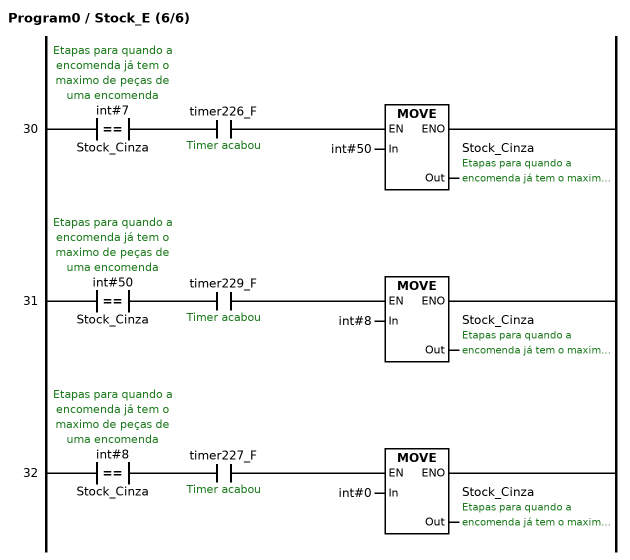
(* [picture p144: Program0 / Stock_E, rungs 30-32] *)
(* Rung 30 *)
IF (int#7 = Stock_Cinza) AND timer226_F THEN Stock_Cinza := int#50; END_IF;
(* Rung 31 *)
IF (int#50 = Stock_Cinza) AND timer229_F THEN Stock_Cinza := int#8; END_IF;
(* Rung 32 *)
IF (int#8 = Stock_Cinza) AND timer227_F THEN Stock_Cinza := int#0; END_IF;

(* Section Stock_S: ladder, written here as Structured Text *)

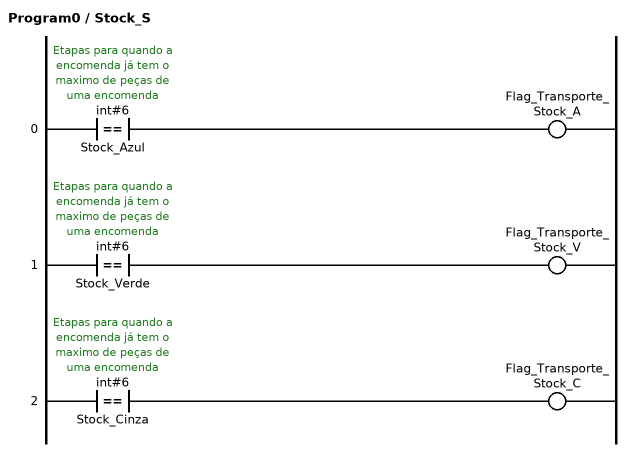
(* Rung 0 *)
Flag_Transporte_Stock_A := int#6 = Stock_Azul;
(* Rung 1 *)
Flag_Transporte_Stock_V := int#6 = Stock_Verde;
(* Rung 2 *)
Flag_Transporte_Stock_C := int#6 = Stock_Cinza;

(* Section Recolhe_Stock_E: ladder, written here as Structured Text *)

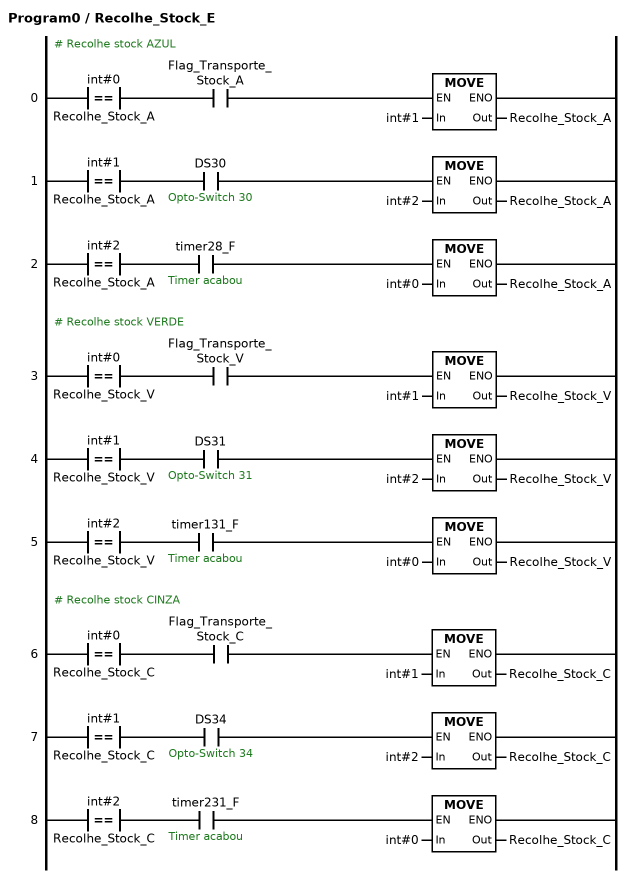
(* Rung 0: # Recolhe stock AZUL *)
IF (int#0 = Recolhe_Stock_A) AND Flag_Transporte_Stock_A THEN Recolhe_Stock_A := int#1; END_IF;
(* Rung 1 *)
IF (int#1 = Recolhe_Stock_A) AND DS30 THEN Recolhe_Stock_A := int#2; END_IF;
(* Rung 2 *)
IF (int#2 = Recolhe_Stock_A) AND timer28_F THEN Recolhe_Stock_A := int#0; END_IF;
(* Rung 3: # Recolhe stock VERDE *)
IF (int#0 = Recolhe_Stock_V) AND Flag_Transporte_Stock_V THEN Recolhe_Stock_V := int#1; END_IF;
(* Rung 4 *)
IF (int#1 = Recolhe_Stock_V) AND DS31 THEN Recolhe_Stock_V := int#2; END_IF;
(* Rung 5 *)
IF (int#2 = Recolhe_Stock_V) AND timer131_F THEN Recolhe_Stock_V := int#0; END_IF;
(* Rung 6: # Recolhe stock CINZA *)
IF (int#0 = Recolhe_Stock_C) AND Flag_Transporte_Stock_C THEN Recolhe_Stock_C := int#1; END_IF;
(* Rung 7 *)
IF (int#1 = Recolhe_Stock_C) AND DS34 THEN Recolhe_Stock_C := int#2; END_IF;
(* Rung 8 *)
IF (int#2 = Recolhe_Stock_C) AND timer231_F THEN Recolhe_Stock_C := int#0; END_IF;

(* Section Recolhe_Stock_S: ladder, written here as Structured Text *)

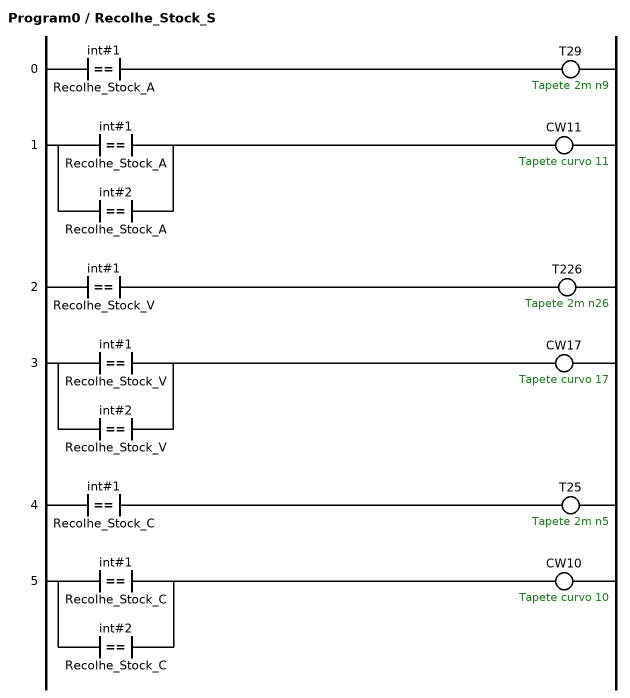
(* Rung 0 *)
T29 := int#1 = Recolhe_Stock_A;
(* Rung 1 *)
CW11 := (int#1 = Recolhe_Stock_A) OR (int#2 = Recolhe_Stock_A);
(* Rung 2 *)
T226 := int#1 = Recolhe_Stock_V;
(* Rung 3 *)
CW17 := (int#1 = Recolhe_Stock_V) OR (int#2 = Recolhe_Stock_V);
(* Rung 4 *)
T25 := int#1 = Recolhe_Stock_C;
(* Rung 5 *)
CW10 := (int#1 = Recolhe_Stock_C) OR (int#2 = Recolhe_Stock_C);

(* Section Recolha_Comum_E: ladder, written here as Structured Text *)

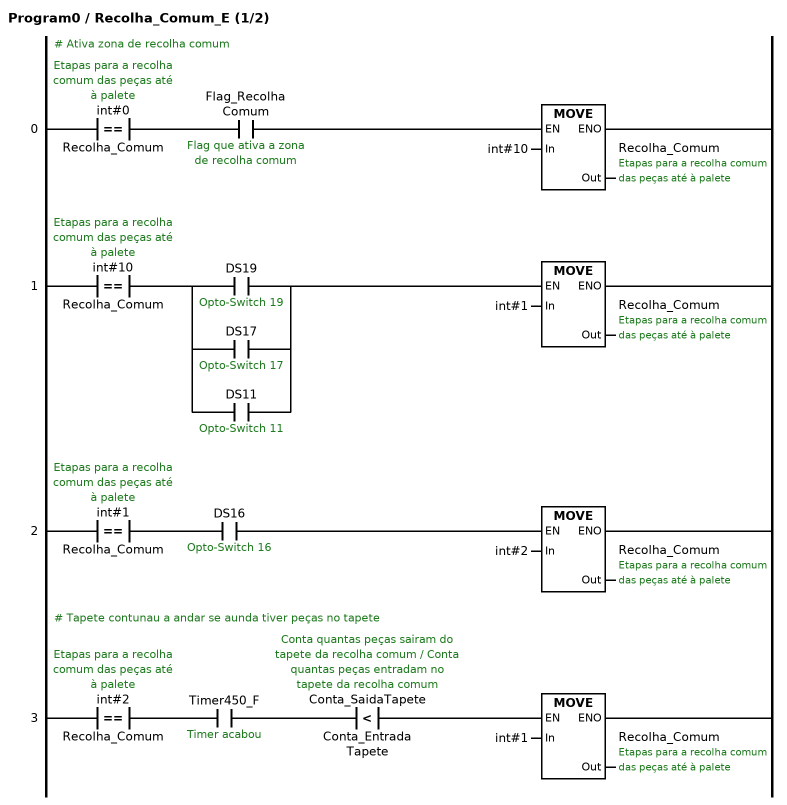
(* Rung 0: # Ativa zona de recolha comum *)
IF (int#0 = Recolha_Comum) AND Flag_RecolhaComum THEN Recolha_Comum := int#10; END_IF;
(* Rung 1 *)
IF (int#10 = Recolha_Comum) AND (DS19 OR DS17 OR DS11) THEN Recolha_Comum := int#1; END_IF;
(* Rung 2 *)
IF (int#1 = Recolha_Comum) AND DS16 THEN Recolha_Comum := int#2; END_IF;
(* Rung 3: # Tapete contunau a andar se aunda tiver peças no tapete *)
IF (int#2 = Recolha_Comum) AND Timer450_F AND (Conta_SaidaTapete < Conta_EntradaTapete) THEN
    Recolha_Comum := int#1;
END_IF;

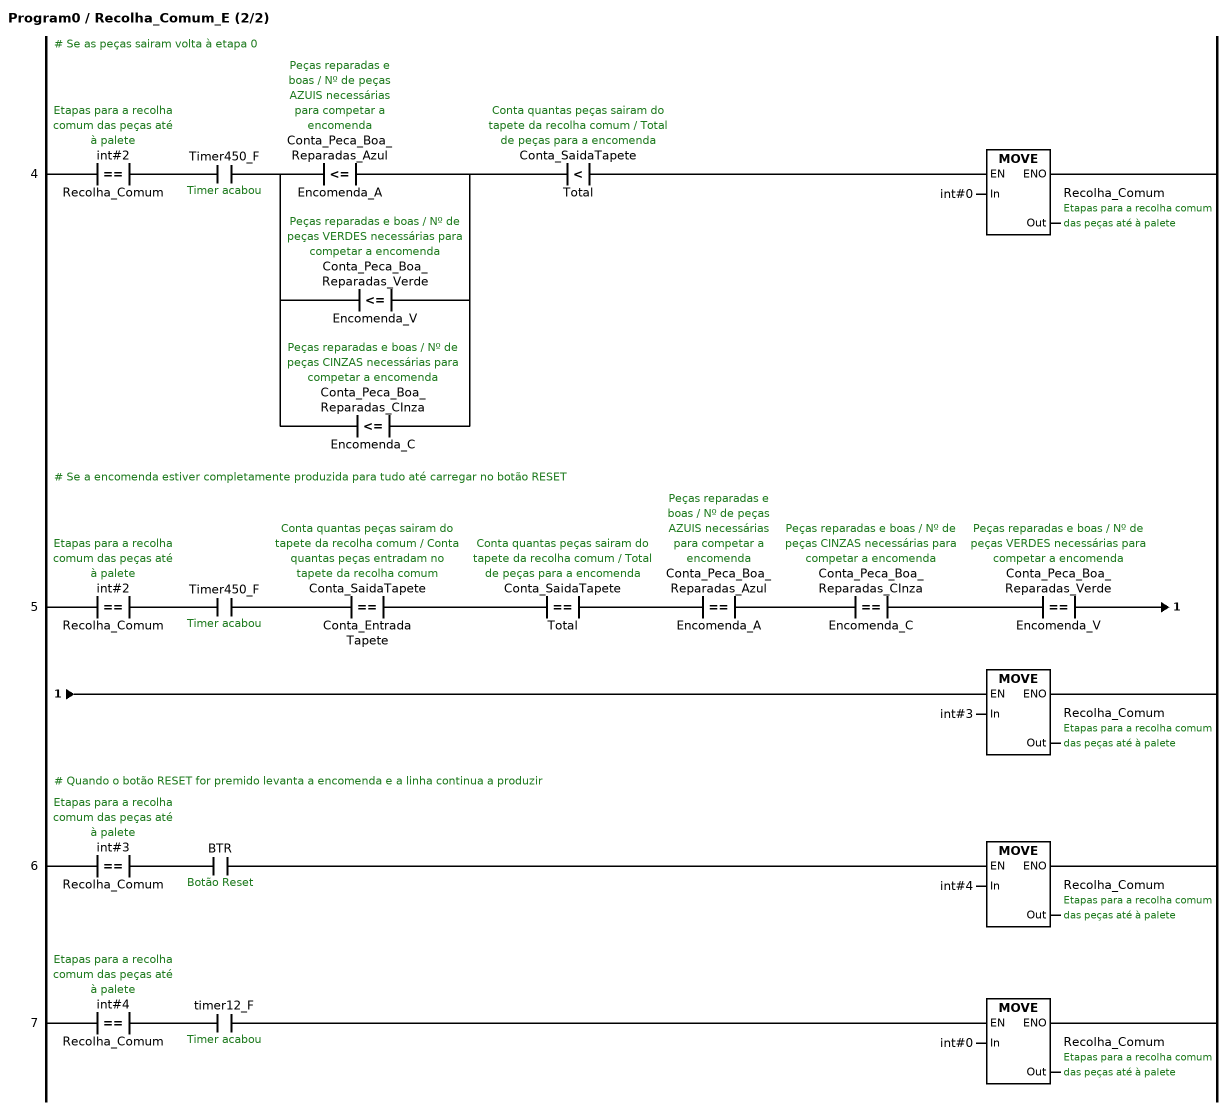
(* Rung 4: # Se as peças sairam volta à etapa 0 *)
IF (int#2 = Recolha_Comum) AND Timer450_F AND ((Conta_Peca_Boa_Reparadas_Azul <= Encomenda_A) OR (Conta_Peca_Boa_Reparadas_Verde <= Encomenda_V) OR (Conta_Peca_Boa_Reparadas_CInza <= Encomenda_C)) AND (Conta_SaidaTapete < Total) THEN
    Recolha_Comum := int#0;
END_IF;
(* Rung 5: # Se a encomenda estiver completamente produzida para tudo até carregar no botão RESET *)
IF (int#2 = Recolha_Comum) AND Timer450_F AND (Conta_SaidaTapete = Conta_EntradaTapete) AND (Conta_SaidaTapete = Total) AND (Conta_Peca_Boa_Reparadas_Azul = Encomenda_A) AND (Conta_Peca_Boa_Reparadas_CInza = Encomenda_C) AND (Conta_Peca_Boa_Reparadas_Verde = Encomenda_V) THEN
    Recolha_Comum := int#3;
END_IF;
(* Rung 6: # Quando o botão RESET for premido levanta a encomenda e a linha continua a produzir *)
IF (int#3 = Recolha_Comum) AND BTR THEN Recolha_Comum := int#4; END_IF;
(* Rung 7 *)
IF (int#4 = Recolha_Comum) AND timer12_F THEN Recolha_Comum := int#0; END_IF;

(* Section Recolha_Comum_S: ladder, written here as Structured Text *)

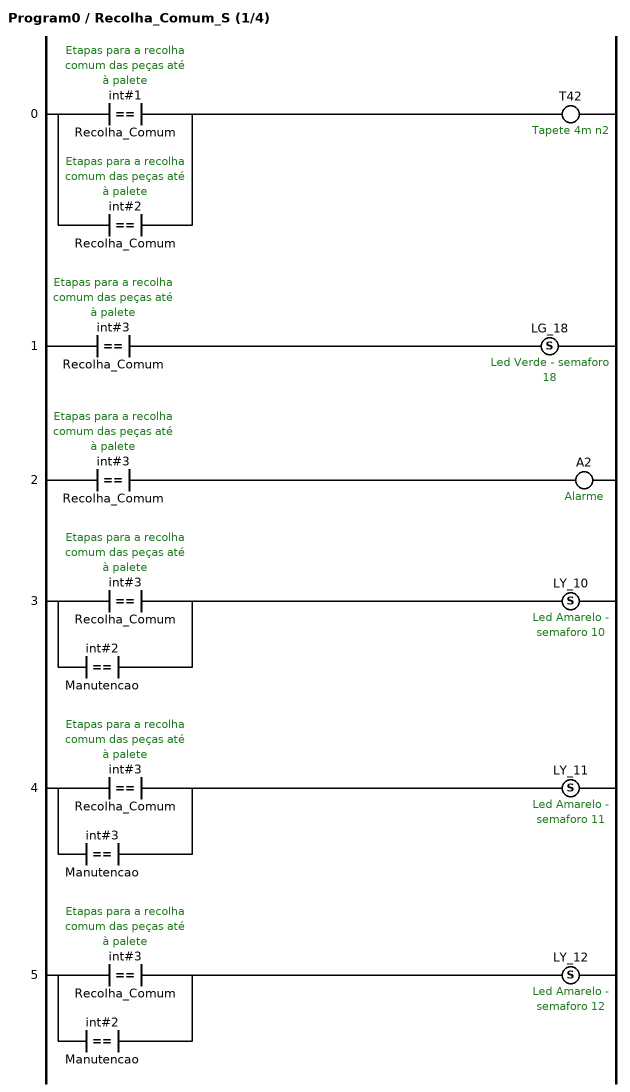
(* Rung 0 *)
T42 := (int#1 = Recolha_Comum) OR (int#2 = Recolha_Comum);
(* Rung 1 *)
IF int#3 = Recolha_Comum THEN LG_18 := TRUE; END_IF;
(* Rung 2 *)
A2 := int#3 = Recolha_Comum;
(* Rung 3 *)
IF (int#3 = Recolha_Comum) OR (int#2 = Manutencao) THEN LY_10 := TRUE; END_IF;
(* Rung 4 *)
IF (int#3 = Recolha_Comum) OR (int#3 = Manutencao) THEN LY_11 := TRUE; END_IF;
(* Rung 5 *)
IF (int#3 = Recolha_Comum) OR (int#2 = Manutencao) THEN LY_12 := TRUE; END_IF;

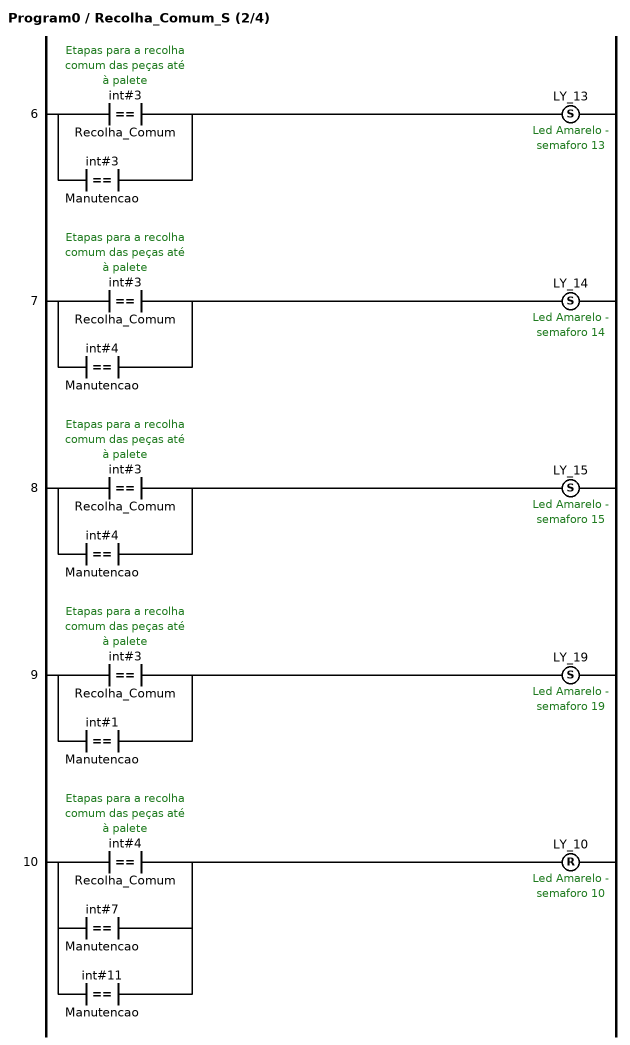
(* Rung 6 *)
IF (int#3 = Recolha_Comum) OR (int#3 = Manutencao) THEN LY_13 := TRUE; END_IF;
(* Rung 7 *)
IF (int#3 = Recolha_Comum) OR (int#4 = Manutencao) THEN LY_14 := TRUE; END_IF;
(* Rung 8 *)
IF (int#3 = Recolha_Comum) OR (int#4 = Manutencao) THEN LY_15 := TRUE; END_IF;
(* Rung 9 *)
IF (int#3 = Recolha_Comum) OR (int#1 = Manutencao) THEN LY_19 := TRUE; END_IF;
(* Rung 10 *)
IF (int#4 = Recolha_Comum) OR (int#7 = Manutencao) OR (int#11 = Manutencao) THEN LY_10 := FALSE; END_IF;

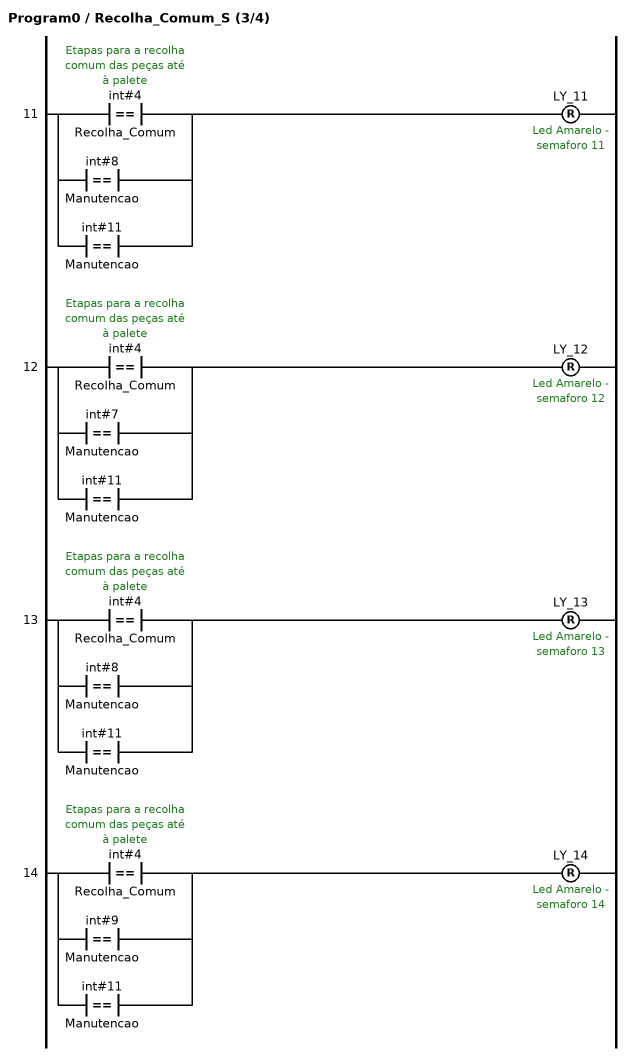
(* Rung 11 *)
IF (int#4 = Recolha_Comum) OR (int#8 = Manutencao) OR (int#11 = Manutencao) THEN LY_11 := FALSE; END_IF;
(* Rung 12 *)
IF (int#4 = Recolha_Comum) OR (int#7 = Manutencao) OR (int#11 = Manutencao) THEN LY_12 := FALSE; END_IF;
(* Rung 13 *)
IF (int#4 = Recolha_Comum) OR (int#8 = Manutencao) OR (int#11 = Manutencao) THEN LY_13 := FALSE; END_IF;
(* Rung 14 *)
IF (int#4 = Recolha_Comum) OR (int#9 = Manutencao) OR (int#11 = Manutencao) THEN LY_14 := FALSE; END_IF;

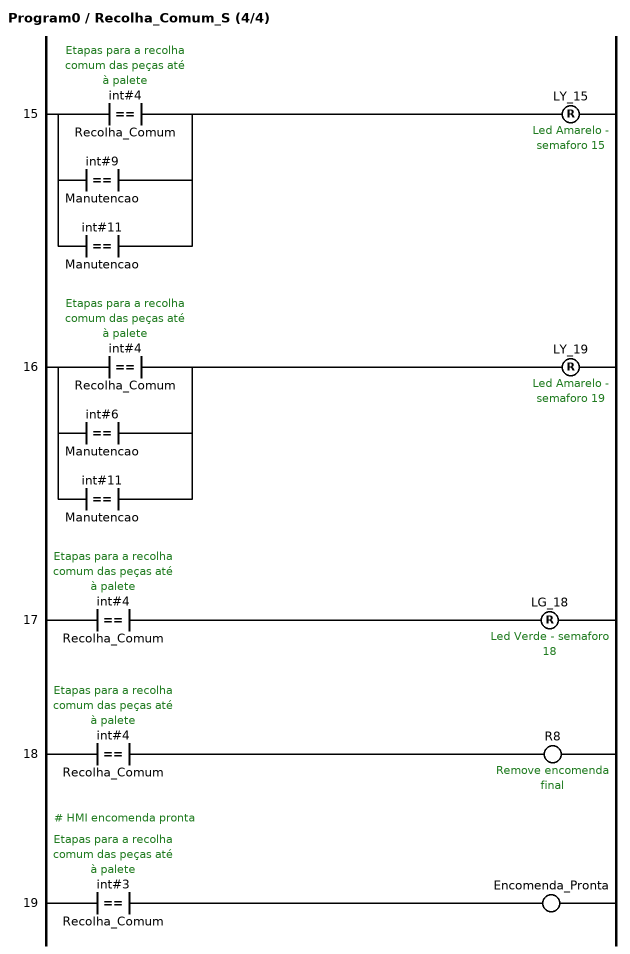
(* Rung 15 *)
IF (int#4 = Recolha_Comum) OR (int#9 = Manutencao) OR (int#11 = Manutencao) THEN LY_15 := FALSE; END_IF;
(* Rung 16 *)
IF (int#4 = Recolha_Comum) OR (int#6 = Manutencao) OR (int#11 = Manutencao) THEN LY_19 := FALSE; END_IF;
(* Rung 17 *)
IF int#4 = Recolha_Comum THEN LG_18 := FALSE; END_IF;
(* Rung 18 *)
R8 := int#4 = Recolha_Comum;
(* Rung 19: # HMI encomenda pronta *)
Encomenda_Pronta := int#3 = Recolha_Comum;
END_PROGRAM

# Device HMI_NA5_0 (NA): not converted